(* IEC 61131-3 sources: rusty/tests/lit/single/enums, 27 files *)

(* ---- enum_ensure_a_combination_of_variables_can_be_assigned_in_function_block.st ---- *)
// RUN: %COMPILE %s && %RUN | %CHECK %s

TYPE EnumType : (
        red,
        green,
        blue
    );
END_TYPE

FUNCTION_BLOCK fb
VAR
    myVar	: EnumType;
END_VAR
VAR_OUTPUT
    outVar	: EnumType;
END_VAR
VAR_IN_OUT
    inOutVar	: EnumType;
END_VAR
myVar := red;
outVar := green;
inOutVar := blue;
END_FUNCTION_BLOCK

PROGRAM prog
VAR
    inOutVar : EnumType;
    outVar: EnumType;
    fb : fb;
END_VAR
    fb(outVar, inOutVar);

    // CHECK: 1
    printf('%d$N', outVar);
    // CHECK: 2
    printf('%d$N', inOutVar);
END_PROGRAM

FUNCTION main
    prog();
END_FUNCTION

(* ---- enum_ensure_in_out_variable_can_be_assigned_in_function_block.st ---- *)
// RUN: %COMPILE %s && %RUN | %CHECK %s

TYPE EnumType : (
        red,
        green,
        blue
    );
END_TYPE

FUNCTION_BLOCK fb
VAR_IN_OUT
    inOutVar	: EnumType;
END_VAR
inOutVar := blue;
END_FUNCTION_BLOCK

PROGRAM prog
VAR
    inOutVar : EnumType;
    fb : fb;
END_VAR
    fb(inOutVar);

    // CHECK: 2
    printf('%d$N', inOutVar);
END_PROGRAM

FUNCTION main
    prog();
END_FUNCTION

(* ---- enum_ensure_output_variable_can_be_assigned_in_function_block.st ---- *)
// RUN: %COMPILE %s && %RUN | %CHECK %s

TYPE EnumType : (
        red,
        green,
        blue
    );
END_TYPE

FUNCTION_BLOCK fb
VAR_OUTPUT
    outVar	: EnumType;
END_VAR
outVar := green;
END_FUNCTION_BLOCK

PROGRAM prog
VAR
    outVar: EnumType;
    fb : fb;
END_VAR
    fb(outVar);

    // CHECK: 1
    printf('%d$N', outVar);
END_PROGRAM

FUNCTION main
    prog();
END_FUNCTION

(* ---- enum_ensure_standard_variable_can_be_assigned_in_function_block.st ---- *)
// RUN: %COMPILE %s && %RUN | %CHECK %s

TYPE EnumType : (
        red,
        green,
        blue
    );
END_TYPE

FUNCTION_BLOCK fb
VAR
    myVar	: EnumType;
END_VAR
myVar := red;
END_FUNCTION_BLOCK

PROGRAM prog
VAR
    fb : fb;
END_VAR
    fb();

    // CHECK: no output
    printf('no output$N');
END_PROGRAM

FUNCTION main
    prog();
END_FUNCTION

(* ---- enum_name_conflicts_with_function_block.st ---- *)
// RUN: %COMPILE %s && %RUN | %CHECK %s

TYPE
    eW : (fooFunc, fooBlock, fooMethod, MyAlias);
END_TYPE

TYPE
    MyAlias : INT;
END_TYPE

FUNCTION fooFunc
    // Does nothing
END_FUNCTION

FUNCTION_BLOCK fooBlock
    METHOD PUBLIC fooMethod
        // Does nothing
    END_METHOD
END_FUNCTION_BLOCK

PROGRAM mainProg
    VAR
        e : eW;
    END_VAR

    // Should be able to assign the enum element to the enum without ambiguity
    e := fooFunc;

    // CHECK: 0
    printf('%d$N', e);

    // Should be able to assign the enum element to the enum without ambiguity
    e := fooBlock;

    // CHECK: 1
    printf('%d$N', e);

    // Should be able to assign the enum element to the enum without ambiguity
    e := fooMethod;

    // CHECK: 2
    printf('%d$N', e);

    // Should be able to assign the enum element to the enum without ambiguity
    e := MyAlias;

    // CHECK: 3
    printf('%d$N', e);

END_PROGRAM

FUNCTION main
    mainProg();
END_FUNCTION

(* ---- debug_enum_explicit_values.st ---- *)
// RUN: %COMPILE_IR %s | %CHECK_IR %s

// Test that enums with explicit values generate correct DIEnumerator entries

TYPE HttpStatus : INT (
    ok := 200,
    not_found := 404,
    server_error := 500
);
END_TYPE

TYPE Powers : DINT (
    one := 1,
    ten := 10,
    hundred := 100,
    thousand := 1000
);
END_TYPE

VAR_GLOBAL
    http_code : HttpStatus := ok;
    power : Powers := one;
END_VAR

PROGRAM prog
    http_code := not_found;
END_PROGRAM

FUNCTION main
    prog();
END_FUNCTION

// CHECK: !DICompositeType(tag: DW_TAG_enumeration_type, name: "HttpStatus"
// CHECK-SAME: elements: ![[HTTP_ELEMENTS:[0-9]+]]

// CHECK: ![[HTTP_ELEMENTS]] = !{![[H0:[0-9]+]], ![[H1:[0-9]+]], ![[H2:[0-9]+]]}
// CHECK: ![[H0]] = !DIEnumerator(name: "ok", value: 200)
// CHECK: ![[H1]] = !DIEnumerator(name: "not_found", value: 404)
// CHECK: ![[H2]] = !DIEnumerator(name: "server_error", value: 500)

// CHECK: !DICompositeType(tag: DW_TAG_enumeration_type, name: "Powers"
// CHECK-SAME: elements: ![[POWER_ELEMENTS:[0-9]+]]

// CHECK: ![[POWER_ELEMENTS]] = !{![[P0:[0-9]+]], ![[P1:[0-9]+]], ![[P2:[0-9]+]], ![[P3:[0-9]+]]}
// CHECK: ![[P0]] = !DIEnumerator(name: "one", value: 1)
// CHECK: ![[P1]] = !DIEnumerator(name: "ten", value: 10)
// CHECK: ![[P2]] = !DIEnumerator(name: "hundred", value: 100)
// CHECK: ![[P3]] = !DIEnumerator(name: "thousand", value: 1000)

(* ---- debug_enum_inline_variables.st ---- *)
// RUN: %COMPILE_IR %s | %CHECK_IR %s

// Test that inline (anonymous) enum variables generate proper debug info
// These are enums declared directly in VAR blocks without TYPE declaration

VAR_GLOBAL
    state : DINT (idle, running, stopped);
    mode : BYTE (manual, automatic);
    priority : INT (low := 1, medium := 5, high := 10);
END_VAR

PROGRAM prog
    state := running;
END_PROGRAM

FUNCTION main
    prog();
END_FUNCTION

// Inline enum for 'state' variable should generate a unique type name
// CHECK: !DICompositeType(tag: DW_TAG_enumeration_type, name: "__global_state"
// CHECK-SAME: baseType: ![[STATE_BASE:[0-9]+]]
// CHECK-SAME: elements: ![[STATE_ELEMENTS:[0-9]+]]

// CHECK: ![[STATE_BASE]] = !DIBasicType(name: "DINT", size: 32, encoding: DW_ATE_signed

// CHECK: ![[STATE_ELEMENTS]] = !{![[S0:[0-9]+]], ![[S1:[0-9]+]], ![[S2:[0-9]+]]}
// CHECK: ![[S0]] = !DIEnumerator(name: "idle", value: 0)
// CHECK: ![[S1]] = !DIEnumerator(name: "running", value: 1)
// CHECK: ![[S2]] = !DIEnumerator(name: "stopped", value: 2)

// Inline enum for 'mode' variable
// CHECK: !DICompositeType(tag: DW_TAG_enumeration_type, name: "__global_mode"
// CHECK-SAME: baseType: ![[MODE_BASE:[0-9]+]]
// CHECK-SAME: size: 8

// CHECK: ![[MODE_BASE]] = !DIBasicType(name: "BYTE", size: 8, encoding: DW_ATE_unsigned

// Inline enum for 'priority' with explicit values
// CHECK: !DICompositeType(tag: DW_TAG_enumeration_type, name: "__global_priority"
// CHECK-SAME: elements: ![[PRIO_ELEMENTS:[0-9]+]]

// CHECK: ![[PRIO_ELEMENTS]] = !{![[PR0:[0-9]+]], ![[PR1:[0-9]+]], ![[PR2:[0-9]+]]}
// CHECK: ![[PR0]] = !DIEnumerator(name: "low", value: 1)
// CHECK: ![[PR1]] = !DIEnumerator(name: "medium", value: 5)
// CHECK: ![[PR2]] = !DIEnumerator(name: "high", value: 10)

(* ---- debug_enum_typed_base_types.st ---- *)
// RUN: %COMPILE_IR %s | %CHECK_IR %s

// Test that typed enums (BYTE, INT, LINT) generate correct debug info with proper base types

TYPE ByteStatus : BYTE (off, on, error);
END_TYPE

TYPE IntLevel : INT (low, medium, high);
END_TYPE

TYPE LintCounter : LINT (zero, one, two);
END_TYPE

VAR_GLOBAL
    status : ByteStatus := off;
    level : IntLevel := low;
    counter : LintCounter := zero;
END_VAR

PROGRAM prog
    status := on;
END_PROGRAM

FUNCTION main
    prog();
END_FUNCTION

// CHECK: !DICompositeType(tag: DW_TAG_enumeration_type, name: "ByteStatus"
// CHECK-SAME: baseType: ![[BYTE_BASE:[0-9]+]]
// CHECK-SAME: size: 8

// CHECK: ![[BYTE_BASE]] = !DIBasicType(name: "BYTE", size: 8, encoding: DW_ATE_unsigned

// CHECK: !DICompositeType(tag: DW_TAG_enumeration_type, name: "IntLevel"
// CHECK-SAME: baseType: ![[INT_BASE:[0-9]+]]
// CHECK-SAME: size: 16

// CHECK: ![[INT_BASE]] = !DIBasicType(name: "INT", size: 16, encoding: DW_ATE_signed

// CHECK: !DICompositeType(tag: DW_TAG_enumeration_type, name: "LintCounter"
// CHECK-SAME: baseType: ![[LINT_BASE:[0-9]+]]
// CHECK-SAME: size: 64

// CHECK: ![[LINT_BASE]] = !DIBasicType(name: "LINT", size: 64, encoding: DW_ATE_signed

(* ---- debug_enum_unsigned_vs_signed.st ---- *)
// RUN: %COMPILE_IR %s | %CHECK_IR %s

// Test that unsigned vs signed enums generate correct isUnsigned flag in DIEnumerator
// Signed types (INT, DINT, LINT) should NOT have isUnsigned flag
// Unsigned types (BYTE, WORD, DWORD, LWORD, UINT, UDINT, ULINT) should have isUnsigned: true

TYPE SignedEnum : INT (neg := -10, zero := 0, pos := 10);
END_TYPE

TYPE UnsignedEnum : BYTE (small, medium, large);
END_TYPE

TYPE DefaultEnum : (a, b, c);  // DINT by default (signed)
END_TYPE

VAR_GLOBAL
    signed_val : SignedEnum := zero;
    unsigned_val : UnsignedEnum := small;
    default_val : DefaultEnum := a;
END_VAR

PROGRAM prog
    signed_val := pos;
END_PROGRAM

FUNCTION main
    prog();
END_FUNCTION

// Signed enum should NOT have isUnsigned flag
// CHECK: !DICompositeType(tag: DW_TAG_enumeration_type, name: "SignedEnum"
// CHECK-SAME: baseType: ![[SIGNED_BASE:[0-9]+]]
// CHECK: ![[SIGNED_BASE]] = !DIBasicType(name: "INT", size: 16, encoding: DW_ATE_signed

// CHECK: !DIEnumerator(name: "neg", value: -10)
// CHECK-NOT: !DIEnumerator(name: "neg", value: -10, isUnsigned: true)
// CHECK: !DIEnumerator(name: "zero", value: 0)
// CHECK-NOT: !DIEnumerator(name: "zero", value: 0, isUnsigned: true)
// CHECK: !DIEnumerator(name: "pos", value: 10)
// CHECK-NOT: !DIEnumerator(name: "pos", value: 10, isUnsigned: true)

// Unsigned enum SHOULD have isUnsigned: true
// CHECK: !DICompositeType(tag: DW_TAG_enumeration_type, name: "UnsignedEnum"
// CHECK-SAME: baseType: ![[UNSIGNED_BASE:[0-9]+]]
// CHECK: ![[UNSIGNED_BASE]] = !DIBasicType(name: "BYTE", size: 8, encoding: DW_ATE_unsigned

// CHECK: !DIEnumerator(name: "small", value: 0, isUnsigned: true)
// CHECK: !DIEnumerator(name: "medium", value: 1, isUnsigned: true)
// CHECK: !DIEnumerator(name: "large", value: 2, isUnsigned: true)

// Default enum (DINT) should NOT have isUnsigned flag
// CHECK: !DICompositeType(tag: DW_TAG_enumeration_type, name: "DefaultEnum"
// CHECK-SAME: baseType: ![[DEFAULT_BASE:[0-9]+]]
// CHECK: ![[DEFAULT_BASE]] = !DIBasicType(name: "DINT", size: 32, encoding: DW_ATE_signed

// CHECK: !DIEnumerator(name: "a", value: 0)
// CHECK-NOT: !DIEnumerator(name: "a", value: 0, isUnsigned: true)

(* ---- debug_enum_variants_not_globals.st ---- *)
// RUN: %COMPILE_IR %s | %CHECK_IR %s

// Test that enum variants are NOT included in global variable debug info
// but the enum type itself and variables using it ARE included
// Variants like Color.red should not appear as global variables

TYPE Color : (red, green, blue);
END_TYPE

TYPE Status : BYTE (inactive, active, error);
END_TYPE

VAR_GLOBAL
    current_color : Color := red;
    current_status : Status := active;
END_VAR

PROGRAM prog
    current_color := green;
END_PROGRAM

FUNCTION main
    prog();
END_FUNCTION

// The global variables should have debug info (in order they appear in IR)
// CHECK: !DIGlobalVariable(name: "current_color"
// CHECK: !DICompositeType(tag: DW_TAG_enumeration_type, name: "Color"
// CHECK: !DIEnumerator(name: "red", value: 0)
// CHECK: !DIEnumerator(name: "green", value: 1)
// CHECK: !DIEnumerator(name: "blue", value: 2)

// CHECK: !DIGlobalVariable(name: "current_status"
// CHECK: !DICompositeType(tag: DW_TAG_enumeration_type, name: "Status"
// CHECK: !DIEnumerator(name: "inactive", value: 0
// CHECK: !DIEnumerator(name: "active", value: 1
// CHECK: !DIEnumerator(name: "error", value: 2

// Enum variants should NOT appear as global variables
// CHECK-NOT: !DIGlobalVariable(name: "red"
// CHECK-NOT: !DIGlobalVariable(name: "green"
// CHECK-NOT: !DIGlobalVariable(name: "blue"
// CHECK-NOT: !DIGlobalVariable(name: "inactive"
// CHECK-NOT: !DIGlobalVariable(name: "active"
// CHECK-NOT: !DIGlobalVariable(name: "error"

(* ---- enum_ensure_a_combination_of_variables_can_be_assigned_in_function.st ---- *)
// RUN: %COMPILE %s && %RUN | %CHECK %s

TYPE EnumType : (
        red,
        green,
        blue
    );
END_TYPE

FUNCTION fn : INT
VAR
    myVar	: EnumType;
END_VAR
VAR_OUTPUT
    outVar	: EnumType;
END_VAR
VAR_IN_OUT
    inOutVar	: EnumType;
END_VAR
myVar := red;
outVar := green;
inOutVar := blue;
END_FUNCTION

PROGRAM prog
VAR
    inOutVar : EnumType;
    outVar: EnumType;
END_VAR
    fn(outVar, inOutVar);

    // CHECK: 1
    printf('%d$N', outVar);
    // CHECK: 2
    printf('%d$N', inOutVar);
END_PROGRAM

FUNCTION main
    prog();
END_FUNCTION

(* ---- enum_ensure_in_out_variable_can_be_assigned_in_function.st ---- *)
// RUN: %COMPILE %s && %RUN | %CHECK %s

TYPE EnumType : (
        red,
        green,
        blue
    );
END_TYPE

FUNCTION fn : INT
VAR_IN_OUT
    inOutVar	: EnumType;
END_VAR
inOutVar := blue;
END_FUNCTION

PROGRAM prog
VAR
    inOutVar : EnumType;
END_VAR
    fn(inOutVar);

    // CHECK: 2
    printf('%d$N', inOutVar);
END_PROGRAM

FUNCTION main
    prog();
END_FUNCTION

(* ---- enum_ensure_output_variable_can_be_assigned_in_function.st ---- *)
// RUN: %COMPILE %s && %RUN | %CHECK %s

TYPE EnumType : (
        red,
        green,
        blue
    );
END_TYPE

FUNCTION fn : INT
VAR_OUTPUT
    outVar	: EnumType;
END_VAR
outVar := green;
END_FUNCTION

PROGRAM prog
VAR
    outVar: EnumType;
END_VAR
    fn(outVar);

    // CHECK: 1
    printf('%d$N', outVar);
END_PROGRAM

FUNCTION main
    prog();
END_FUNCTION

(* ---- enum_ensure_pointer_to_pointer_can_be_assigned.st ---- *)
// RUN: %COMPILE %s && %RUN | %CHECK %s

VAR_GLOBAL
    someEnum : EnumType;
END_VAR

TYPE EnumType : (
        red,
        green,
        blue
    );
END_TYPE

FUNCTION fn : INT
VAR_IN_OUT
    myVar	: EnumType;
END_VAR
myVar := green;
END_FUNCTION

PROGRAM prog
VAR
    enumRef : reference to EnumType ref= someEnum;
END_VAR
    fn(enumRef);

    // CHECK: 1
    printf('%d$N', enumRef);
END_PROGRAM

FUNCTION main
    prog();
END_FUNCTION

(* ---- enum_ensure_standard_variable_can_be_assigned_in_function.st ---- *)
// RUN: %COMPILE %s && %RUN | %CHECK %s

TYPE EnumType : (
        red,
        green,
        blue
    );
END_TYPE

FUNCTION fn : INT
VAR
    myVar	: EnumType;
END_VAR
myVar := red;
END_FUNCTION

PROGRAM prog
    fn();

    // CHECK: no output
    printf('no output$N');
END_PROGRAM

FUNCTION main
    prog();
END_FUNCTION

(* ---- enum_ensure_zero_variant_initializer_works_with_constant_variables.st ---- *)
// RUN: %COMPILE %s && %RUN | %CHECK %s

VAR_GLOBAL CONSTANT
    MYCONST: INT := 0;
END_VAR

// Test enum with no explicit default and a zero variant that is NOT also the first variant - BUT instead of a literal use a constant to initialize
TYPE Status : INT (
    active := 1,
    inactive := MYCONST,
    error := 2
);
END_TYPE

VAR_GLOBAL
    s_global: Status;  // Should initialize to inactive
END_VAR

PROGRAM prog
VAR
    s1 : Status;  // Should initialize to inactive
END_VAR
    // CHECK: 0
    printf('%d$N', s1);  // inactive

    // CHECK: 0
    printf('%d$N', s_global);  // inactive
END_PROGRAM

FUNCTION main
    prog();
END_FUNCTION

(* ---- hwmap_enum_no_stack_overflow.st ---- *)
// --hwmap-file must not stack-overflow on programs that
// contain enum typed variables. The instance iterator used to descend into
// enum variants, re-entering the same enum type forever until the stack
// was exhausted.

// First we make sure that the hwmap file does not stack overflow
// RUN: timeout 10s %PLC -i %UTILS --check --hwmap-file=%t.hwmap.json %s

// Then we do a sanity run to make sure the program executes to completion and produces the expected output
// RUN: %COMPILE %s && %RUN | %CHECK %s

TYPE enumType : (
    element0,
    element1
);
END_TYPE

VAR_GLOBAL
    myGlobalEnum : enumType;
END_VAR

PROGRAM mainProg
VAR
    myLocalEnum : enumType;
END_VAR
END_PROGRAM

FUNCTION main
    mainProg();

    // CHECK: Complete
    printf('Complete$N');
END_FUNCTION

(* ---- typed_enum_61131_syntax_with_default.st ---- *)
// RUN: %COMPILE %s && %RUN | %CHECK %s

// Test IEC 61131-3 syntax: TYPE NAME : TYPE (variants) := default;
TYPE Status : DWORD (
    inactive := 16#00000000,
    active := 16#00000001,
    error := 16#FFFFFFFF
) := inactive;
END_TYPE

VAR_GLOBAL
    s_global: Status;  // Should initialize to inactive (explicit default)
END_VAR

PROGRAM prog
VAR
    s1 : Status;  // Should initialize to inactive (explicit default)
    s2 : Status := active;
    s3 : Status := error;
END_VAR
    // CHECK: 0
    printf('%d$N', s1);  // inactive (default)

    // CHECK: 1
    printf('%d$N', s2);  // active

    // CHECK: -1
    printf('%d$N', s3);  // error (as signed)

    // CHECK: 0
    printf('%d$N', s_global);  // inactive (default)
END_PROGRAM

FUNCTION main
    prog();
END_FUNCTION

(* ---- typed_enum_byte_values_are_correct.st ---- *)
// RUN: %COMPILE %s && %RUN | %CHECK %s

// Test BYTE enum values work correctly
TYPE Status : BYTE (inactive := 0, active := 1, error := 255);
END_TYPE

VAR_GLOBAL
    status_global: Status := active;
END_VAR

PROGRAM prog
VAR
    s1 : Status := inactive;
    s2 : Status := active;
    s3 : Status := error;
END_VAR
    // CHECK: 0
    printf('%d$N', s1);  // inactive

    // CHECK: 1
    printf('%d$N', s2);  // active

    // CHECK: 255
    printf('%d$N', s3);  // error

    // CHECK: 1
    printf('%d$N', status_global);  // active
END_PROGRAM

FUNCTION main
    prog();
END_FUNCTION

(* ---- typed_enum_codesys_syntax_with_default.st ---- *)
// RUN: %COMPILE %s && %RUN | %CHECK %s

// Test Codesys syntax: TYPE NAME : (variants) TYPE := default;
TYPE Priority : (
    low := 10,
    medium := 20,
    high := 30
) INT := medium;
END_TYPE

VAR_GLOBAL
    p_global: Priority;  // Should initialize to medium (explicit default)
END_VAR

PROGRAM prog
VAR
    p1 : Priority;  // Should initialize to medium (explicit default)
    p2 : Priority := high;
END_VAR
    // CHECK: 20
    printf('%d$N', p1);  // medium (default)

    // CHECK: 30
    printf('%d$N', p2);  // high

    // CHECK: 20
    printf('%d$N', p_global);  // medium (default)
END_PROGRAM

FUNCTION main
    prog();
END_FUNCTION

(* ---- typed_enum_initialized_with_typed_literal.st ---- *)
// RUN: %COMPILE %s && %RUN | %CHECK %s
PROGRAM mainProg
    foo();
END_PROGRAM

FUNCTION foo
    VAR
        vEnum : myEnum := e2;
    END_VAR

    printf('%d$N', vEnum);

END_FUNCTION

TYPE
	myEnum : (e1, e2:=BYTE#30) BYTE;
END_TYPE

FUNCTION main
    // CHECK: 30
    mainProg();
END_FUNCTION

(* ---- typed_enum_initialized_with_typed_literal_with_no_intermediate_function.st ---- *)
// RUN: %COMPILE %s && %RUN | %CHECK %s
PROGRAM mainProg
    VAR
        vEnum : myEnum := e2;
    END_VAR

    printf('%d$N', vEnum);
END_PROGRAM

TYPE
	myEnum : (e1, e2:=BYTE#30) BYTE;
END_TYPE

FUNCTION main
    // CHECK: 30
    mainProg();
END_FUNCTION

(* ---- typed_enum_various_integer_types.st ---- *)
// RUN: %COMPILE %s && %RUN | %CHECK %s

// Test various integer types work correctly
TYPE ByteEnum : BYTE (a := 1, b := 2);
END_TYPE

TYPE IntEnum : INT (x := 100, y := 200);
END_TYPE

TYPE DwordEnum : DWORD (big := 16#FFFF0000, small := 16#00000000);
END_TYPE

TYPE LintEnum : LINT (huge := 9223372036854775807, semi_huge := 123421341234);  // Max LINT
END_TYPE

PROGRAM prog
VAR
    be : ByteEnum := b;
    ie : IntEnum := y;
    de : DwordEnum := big;
    le : LintEnum := huge;
END_VAR
    // CHECK: 2
    printf('%d$N', be);  // BYTE

    // CHECK: 200
    printf('%d$N', ie);  // INT

    // CHECK: -65536
    printf('%d$N', de);  // DWORD (as signed)

    // CHECK: 9223372036854775807
    printf('%lld$N', le);  // LINT
END_PROGRAM

FUNCTION main
    prog();
END_FUNCTION

(* ---- typed_enum_with_zero_and_explicit_default.st ---- *)
// RUN: %COMPILE %s && %RUN | %CHECK %s

// Test enum with zero variant BUT explicit default - should use explicit default
TYPE Status : INT (
    inactive := 0,
    active := 1,
    error := 2
) := active;
END_TYPE

VAR_GLOBAL
    s_global: Status;  // Should initialize to active (explicit default)
END_VAR

PROGRAM prog
VAR
    s1 : Status;  // Should initialize to active (explicit default), not inactive
    s2 : Status := error;
END_VAR
    // CHECK: 1
    printf('%d$N', s1);  // active (explicit default overrides zero)

    // CHECK: 2
    printf('%d$N', s2);  // error

    // CHECK: 1
    printf('%d$N', s_global);  // active (explicit default)
END_PROGRAM

FUNCTION main
    prog();
END_FUNCTION

(* ---- typed_enum_with_zero_no_default.st ---- *)
// RUN: %COMPILE %s && %RUN | %CHECK %s

// Test enum with zero variant and NO explicit default - should init to zero
TYPE Status : INT (
    inactive := 0,
    active := 1,
    error := 2
);
END_TYPE

VAR_GLOBAL
    s_global: Status;  // Should initialize to inactive (zero value)
END_VAR

PROGRAM prog
VAR
    s1 : Status;  // Should initialize to inactive (zero value)
    s2 : Status := active;
END_VAR
    // CHECK: 0
    printf('%d$N', s1);  // inactive (zero default)

    // CHECK: 1
    printf('%d$N', s2);  // active

    // CHECK: 0
    printf('%d$N', s_global);  // inactive (zero default)
END_PROGRAM

FUNCTION main
    prog();
END_FUNCTION

(* ---- typed_enum_without_zero_no_default.st ---- *)
// RUN: %COMPILE %s && %RUN | %CHECK %s

// Test enum without zero variant and NO explicit default - should init to first element
TYPE Priority : INT (
    low := 10,
    medium := 20,
    high := 30
);
END_TYPE

VAR_GLOBAL
    p_global: Priority;  // Should initialize to low (first element)
END_VAR

PROGRAM prog
VAR
    p1 : Priority;  // Should initialize to low (first element)
    p2 : Priority := high;
END_VAR
    // CHECK: 10
    printf('%d$N', p1);  // low (first element default)

    // CHECK: 30
    printf('%d$N', p2);  // high

    // CHECK: 10
    printf('%d$N', p_global);  // low (first element default)
END_PROGRAM

FUNCTION main
    prog();
END_FUNCTION

(* ---- typed_enum_without_zero_with_default.st ---- *)
// RUN: %COMPILE %s && %RUN | %CHECK %s

// Test enum without zero variant but WITH explicit default - should init to explicit default
TYPE PRIORITY : INT (
    low := 10,
    medium := 20,
    high := 30
) := medium;
END_TYPE

VAR_GLOBAL
    p_global: PRIORITY;
END_VAR

PROGRAM prog
VAR
    p1 : PRIORITY;  // Should initialize to medium (explicit default), not low
    p2 : PRIORITY := high;
END_VAR
    // CHECK: 20
    printf('%d$N', p1);  // Should be medium (explicit default)

    // CHECK: 30
    printf('%d$N', p2);  // high

    p1 := PRIORITY.low;
    // CHECK: 10
    printf('%d$N', p1);  // low

    // CHECK: 20
    printf('%d$N', p_global); // medium
END_PROGRAM

FUNCTION main
    prog();
END_FUNCTION
